TYPE ST_SafeOut_PlcIn :
STRUCT
	ES1_PB_State	:BOOL;
	ES2_PB_State	:BOOL;
	ES3_PB1_State	:BOOL;
	ES3_PB2_State	:BOOL;
	ES4_PB_State	:BOOL;
	
	ES1_State		: BOOL;
	ES2_State		: BOOL;
	ES3_State		: BOOL;
	ES4_State		: BOOL;
	
	TankLocked_CIP_T91: BOOL;
	TankLocked_CIP_T92: BOOL;
	TankLocked_CIP_T93: BOOL;
	TankLocked_CIP_T94: BOOL;
	TankLocked_Marinade_T1: BOOL;
	TankLocked_Marinade_T2: BOOL;
	TankLocked_Color_T3: BOOL;
	TankLocked_Color_T4: BOOL;

END_STRUCT
END_TYPE

(* stored: Version 1.1.0.1, ProductVersion 3.1.4024.13
   DUT ST_SafeOut_PlcIn: Id {6945b16e-45f5-45f1-ba6e-89c09d6c8d7f} *)
